{attribute 'qualified_only'}
VAR_GLOBAL
    config : ST_ConveyorConfig;
    running : ARRAY[1..3] OF BOOL;
    actualSpeed : ARRAY[1..3] OF LREAL;
END_VAR

(* stored: Version 1.1.0.1, ProductVersion 3.1 *)
